Fanuc KAREL source: KT00326.KL

PROGRAM KT00326
%NOLOCKGROUP
VAR
  P1: JOINTPOS
  P2: JOINTPOS
  OUT: BOOLEAN
BEGIN
  OUT = P1 <> P2
END KT00326
